ABB RobotStudio station: TPL1_Heredia_Biancuzzo.rspag

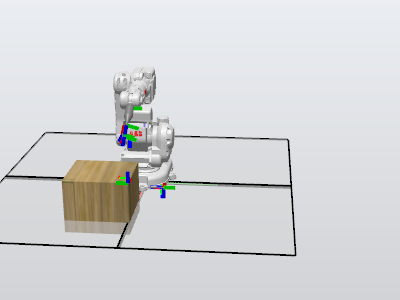
--- station ---
Station TPL1 (saved by RobotStudio 25.5.11605.0)
Controller IRB140_6_81
  mechanical unit ROB_1: IRB140_6_81_C_03, 6 joints, base frame (0, 0, 0) mm
Layout (positions relative to the parent item):
  - IRB140_6_81_C_03 [mechanism, from %ABB.RobotStudio.Models.IRB140%\IRB140_6_81_C_G_03.rslib] at (0, 0, 0) mm; joint values [0, 0, 0, 0, 0.5236, 0] (rad or m)
  - Mesa [part], size 365 x 405 x 340 mm
  - Perno [part] at (904.35, 122.3, 711.04) mm, size 20 x 100 x 20 mm
  - Pinza [mechanism] at (506.29, 0, 679.5) mm, rotated rx 180 ry 60 rz 180 deg
      TCP Pinza at (0, 0, 137) mm, rotated rx 0 ry 0 rz -22.5 deg
      links: Dummy
Attachment: Pinza is attached to IRB140_6_81_C_03 / Link6
EventTableEntry 2362: ActivationMode=2, Cyclic=false, Group=, Trigger=DO_Pinza 2363, Actions=[EventTableActionAttach 2364], Comment=
EventTableTriggerIO 2363: Operator=0, IOValue=[1], IRC5Controller=? -1, SignalSource=IRB140_6_81 1261
EventTableActionAttach 2364: MountObject=false, FlangeIndext=0, FindNearest=false, AttachmentParent=Pinza 2358, AttachmentChild=Perno 2354, Offset=[X=1, Y=0, Z=0, W=0, X=0, Y=1, Z=0, W=0, X=0, Y=0, Z=1, W=0, X=0, Y=0, Z=0, W=1]
EventTableEntry 2365: ActivationMode=2, Cyclic=false, Group=, Trigger=DO_Pinza 2366, Actions=[EventTableActionDetach 2367], Comment=
EventTableTriggerIO 2366: Operator=0, IOValue=[0], IRC5Controller=? -1, SignalSource=IRB140_6_81 1261
EventTableActionDetach 2367: AttachmentParent=Pinza 2358, AttachmentChild=Perno 2354
Collision set Conjunto de colisión_1: Mesa against Perno, IRB140_6_81_C_03, Pinza, near miss 0.01 m
Targets, tools, work objects and paths stored in the station and not in the controller backup, written as RAPID:
! task T_ROB1
MODULE Module1
  PERS tooldata PinzaPerno:=[TRUE,[[83.1492,-34.4415,137],[0.69352,0.13795,0.69352,-0.13795]],[0.5,[0,0,100],[1,0,0,0],0,0,0]];
  PROC Path()
    MoveJ Home,v50,z100,Pinza\WObj:=Terna_Origen;
    AbrirPinza;
    MoveJ Offs(Pick, 0, 0, OffsetPick),v100,z100,Pinza\WObj:=Terna_Dispenser;
    MoveL Pick,v10,fine,Pinza\WObj:=Terna_Dispenser;
    CerrarPinza;
    MoveL Offs(Pick, 0, 0, OffsetPick),v10,z100,Pinza\WObj:=Terna_Dispenser;
    MoveJ Offs(Place, 0, 0, OffsetPlace),v100,z100,PinzaPerno\WObj:=Terna_Mesa;
    MoveL Offs(Place, 0, 0, OffsetHole),v10,fine,PinzaPerno\WObj:=Terna_Mesa;
    AbrirPinza;
    MoveL Offs(Place, 0, 0, OffsetPlace),v10,z100,PinzaPerno\WObj:=Terna_Mesa;
    MoveJ Home,v50,z100,Pinza\WObj:=Terna_Origen;
  ENDPROC
ENDMODULE


--- Controller Data/IRB140_6_81/RAPID/TASK1/PROGMOD/CalibData.mod ---
MODULE CalibData
    PERS tooldata Pinza:=[TRUE,[[0,0,137],[0.980785,0,0,-0.19509]],[0.5,[0,0,100],[1,0,0,0],0,0,0]];
    PERS tooldata PinzaPernoLateral := [TRUE,[[0,0,227],[0.980785,0,0,-0.19509]],[0.5,[0,0,100],[1,0,0,0],0,0,0]];
    PERS tooldata PinzaPernoVertical := [TRUE,[[83.1492,-34.4415,137],[0.69352,0.13795,0.69352,-0.13795]],[0.5,[0,0,100],[1,0,0,0],0,0,0]];
    PERS wobjdata Terna_Origen:=[FALSE,TRUE,"",[[0,0,0],[0,0,0,1]],[[0,0,0],[1,0,0,0]]];
    PERS wobjdata Terna_Mesa:=[FALSE,TRUE,"",[[665,5,260],[0,0,0,1]],[[0,0,0],[1,0,0,0]]];
    PERS wobjdata Terna_Dispenser:=[FALSE,TRUE,"",[[400,180,130],[0,0,1,0]],[[0,0,0],[1,0,0,0]]];
ENDMODULE

--- Controller Data/IRB140_6_81/RAPID/TASK1/PROGMOD/Module1.mod ---
MODULE Module1
    CONST robtarget Home:=[[-500,7.461,500],[0,0,1,0],[-1,0,-2,0],[9E+09,9E+09,9E+09,9E+09,9E+09,9E+09]];
    CONST robtarget Place:=[[65,65,0],[0,1,0,0],[-1,0,-2,0],[9E+09,9E+09,9E+09,9E+09,9E+09,9E+09]];
    CONST robtarget PickVertical:=[[0,-10,0],[0.707106781,0,0,-0.707106781],[0,0,0,0],[9E+09,9E+09,9E+09,9E+09,9E+09,9E+09]];
    CONST robtarget PickLateral:=[[0,-10,0],[0.707106781,0.707106781,0,0],[0,0,0,0],[9E+09,9E+09,9E+09,9E+09,9E+09,9E+09]];

    CONST intnum TiempoHerramienta := 5;
    CONST intnum OffsetPick := -100;
    CONST intnum OffsetPlace := 150;
    CONST intnum OffsetHole := -15;
    CONST intnum Conf := 0;

    CONST speeddata VMax := v30;
    CONST speeddata VMin := v10;

    VAR pose PosePinzaPernoLateral;
    VAR pose PosePinzaPernoVertical;

    !***********************************************************
    ! Autor: rocio
    !***********************************************************

    PROC main()
        IF Conf = 1 THEN
            PosePinzaPernoLateral := PoseMult(Pinza.tframe, [[0,0,90],[1,0,0,0]]);
            PinzaPernoLateral:=[TRUE,PosePinzaPernoLateral,[0.5,[0,0,100],[1,0,0,0],0,0,0]];
            Path PinzaPernoLateral, PickLateral;
        ELSE
            PosePinzaPernoVertical := PoseMult(Pinza.tframe, [[90,0,0],[0.7071,0,0.7071,0]]);
            PinzaPernoVertical:=[TRUE,PosePinzaPernoVertical,[0.5,[0,0,100],[1,0,0,0],0,0,0]];
            Path PinzaPernoVertical, PickVertical;
        ENDIF

    ENDPROC
    PROC Path (PERS tooldata PinzaPerno, robtarget Pick)
        MoveJ Home,VMax,fine,Pinza\WObj:=Terna_Origen;
        AbrirPinza;

        MoveJ Offs(Pick, 0, 0, OffsetPick),VMax,z100,Pinza\WObj:=Terna_Dispenser;
        MoveL Pick,VMin,fine,Pinza\WObj:=Terna_Dispenser;
        CerrarPinza;
        MoveL Offs(Pick, 0, 0, OffsetPick),VMin,z100,Pinza\WObj:=Terna_Dispenser;

        MoveJ Offs(Place, 0, 0, OffsetPlace),VMax,z100,PinzaPerno\WObj:=Terna_Mesa;
        MoveL Offs(Place, 0, 0, OffsetHole),VMin,fine,PinzaPerno\WObj:=Terna_Mesa;
        AbrirPinza;
        MoveL Offs(Place, 0, 0, OffsetPlace),VMin,fine,PinzaPerno\WObj:=Terna_Mesa;

        MoveJ Home,VMax,fine,Pinza\WObj:=Terna_Origen;
    ENDPROC

    PROC AbrirPinza()
        SetDO DO_Pinza, 0;
        WaitTime TiempoHerramienta;
    ENDPROC
    PROC CerrarPinza()
        SetDO DO_Pinza, 1;
        WaitTime TiempoHerramienta;
    ENDPROC
ENDMODULE

--- Controller Data/IRB140_6_81/SYSPAR/EIO.cfg ---
EIO:CFG_1.0:6:1::
#
EIO_SIGNAL:

      -Name "DO_Pinza" -SignalType "DO" -Access "All"
